Staubli VAL3: lifebit.pgx

public program lifebit()
begin
  //  _nClock=0
  //  do
  if clock()-_nClock>1
    _nClock=clock()
    bLifebit=!bLifebit
  endIf


  //  delay(0)
  //  until false
end
